Staubli VAL3: Prog_Name_Tha.pjx

--- Prog_Name_Tha.pjx ---
Parameters version=s7.5.3 stackSize=5000 millimeterUnit=true
Program file=MoveJoint.pgx
Program file=MoveLine.pgx
Program file=start.pgx
Program file=stop.pgx
Program file=main.pgx
Data file=Prog_Name_Tha.dtx

--- Prog_Name_Tha.dtx ---
mdesc mNomSpeed
frame fFrame1 = {x=250.000, y=300.000, z=-10.000, rx=-0.000, ry=0.000, rz=90.000, fatherId=world[0]}
dio Input[16]
  [0] = {link=BasicIO-1\%I0}
  [1] = {link=BasicIO-1\%I1}
  [2] = {link=BasicIO-1\%I2}
  [3] = {link=BasicIO-1\%I3}
  [4] = {link=BasicIO-1\%I4}
  [5] = {link=BasicIO-1\%I5}
  [6] = {link=BasicIO-1\%I6}
  [7] = {link=BasicIO-1\%I7}
  [8] = {link=BasicIO-1\%I8}
  [9] = {link=BasicIO-1\%I9}
  [10] = {link=BasicIO-1\%I10}
  [11] = {link=BasicIO-1\%I11}
  [12] = {link=BasicIO-1\%I12}
  [13] = {link=BasicIO-1\%I13}
  [14] = {link=BasicIO-1\%I14}
  [15] = {link=BasicIO-1\%I15}
dio Output[16]
  [0] = {link=BasicIO-1\%Q0}
  [1] = {link=BasicIO-1\%Q1}
  [2] = {link=BasicIO-1\%Q2}
  [3] = {link=BasicIO-1\%Q3}
  [4] = {link=BasicIO-1\%Q4}
  [5] = {link=BasicIO-1\%Q5}
  [6] = {link=BasicIO-1\%Q6}
  [7] = {link=BasicIO-1\%Q7}
  [8] = {link=BasicIO-1\%Q8}
  [9] = {link=BasicIO-1\%Q9}
  [10] = {link=BasicIO-1\%Q10}
  [11] = {link=BasicIO-1\%Q11}
  [12] = {link=BasicIO-1\%Q12}
  [13] = {link=BasicIO-1\%Q13}
  [14] = {link=BasicIO-1\%Q14}
  [15] = {link=BasicIO-1\%Q15}
tool tCurrentTool = {x=10.000, y=0.000, z=120.000, rx=-0.000, ry=15.000, rz=-0.000, fatherId=flange[0], ioLink=ValveIO/valve1}
mdesc mCurrentSpeed
pointRx pPointRx = {fatherId=fFrame1[0]}
pointRx pPointRx2 = {fatherId=fFrame1[0]}

--- main.pgx ---
program main()
begin
  close(tCurrentTool)
  pPointRx.config.shoulder = lefty
  pPointRx.config.elbow = epositive
  pPointRx.config.wrist = wpositive
  pPointRx2.config.shoulder = lefty
  pPointRx2.config.elbow = epositive
  pPointRx2.config.wrist = wpositive
  mCurrentSpeed.tvel = 100.00
  mCurrentSpeed.blend = joint
  mCurrentSpeed.reach = 0.010
  mCurrentSpeed.leave = 0.010
  // Program Prog_Name_That_Is_Very_Long_123 start
  // Program generated by VerticalBot Studio for Staubli RX160 on 25/10/2026 12:00:00
  // Using nominal kinematics.
  mCurrentSpeed.tvel = 1000.000
  mCurrentSpeed.reach = 10.000
  mCurrentSpeed.leave = 10.000
  call MoveJoint(10.00000,20.00000,90.00000,30.00000,45.00000,60.00000)
  call MoveLine(1077.300,-56.172,837.243,-146.156,25.288,-102.118)
  mCurrentSpeed.reach = 0.500
  mCurrentSpeed.leave = 0.500
  call MoveLine(1005.190,-118.362,847.372,-147.806,26.655,-97.799)
  delay(0.000)
  delay(1.500)
  popUpMsg("Say "hi" to the operator")
  // A long comment line that exceeds the usual controller limits for comments by far, really
  Output[12]=false
  OUT_A=true
  watch(Input[4]==false,1000.0)
  watch(IN_B==true)
  //call prog:Program_With_A_Long_Name_ABCDEFGHIJ()
  call MoveLine(1077.300,-56.172,837.243,-146.156,25.288,-102.118)
  mCurrentSpeed.reach = -1.000
  mCurrentSpeed.leave = -1.000
  call MoveJoint(10.00000,20.00000,90.00000,30.00000,45.00000,60.00000)

  waitEndMove()
  // Program Prog_Name_That_Is_Very_Long_123 end

end

--- start.pgx ---
program start()
begin
  call main()
end

--- MoveJoint.pgx ---
program MoveJoint(num x_nJ1, num x_nJ2, num x_nJ3, num x_nJ4, num x_nJ5, num x_nJ6)
  local joint l_jJoint
begin
  l_jJoint.j1 = x_nJ1
  l_jJoint.j2 = x_nJ2
  l_jJoint.j3 = x_nJ3
  l_jJoint.j4 = x_nJ4
  l_jJoint.j5 = x_nJ5
  l_jJoint.j6 = x_nJ6
  movej(l_jJoint,tCurrentTool ,mCurrentSpeed)
end

--- MoveLine.pgx ---
program MoveLine(num x_nX, num x_nY, num x_nZ, num x_nRx, num x_nRy, num x_nRz)
begin
  pPointRx.trsf.x = x_nX
  pPointRx.trsf.y = x_nY
  pPointRx.trsf.z = x_nZ
  pPointRx.trsf.rx = x_nRx
  pPointRx.trsf.ry = x_nRy
  pPointRx.trsf.rz = x_nRz
  movel(pPointRx,tCurrentTool,mCurrentSpeed)
end

--- stop.pgx ---
program stop()
begin
end
